(* IEC 61131-3 sources: IEC61131-3_ST_SCL_Mutation_Generator/Tests/mutatedCode_pressure_sensors_m, 18 files *)

(* ---- M1405.st ---- *)
FUNCTION_BLOCK "MAIN"
{ S7_Optimized_Access := 'FALSE' }
VERSION : 1.0

VAR_OUTPUT
    Done : Bool;              // TRUE when the operation has completed
END_VAR

VAR
    presure_sensor : UInt := 10;
    temp_sensor : Int := 2;
    relay : Bool := TRUE;
    counter : UInt;
    error_code : Int;
    error : Bool := TRUE;
    GT1_OUT : Bool;
END_VAR

BEGIN

    // IEC "PROGRAM MAIN" implemented as an SCL function block so it can be
    // instantiated and verified (properties refer to instance.<variable>).

    #Done := FALSE;

    // Loop through the pressure sensor samples
    #counter := 0;
    WHILE #counter > #presure_sensor DO (* MUTATED: REL_OP_REPLACE *)

        #counter := #counter + 1;

        // Adjust the temperature sensor value, with overflow protection
        IF #temp_sensor < 32767 THEN
            #temp_sensor := #temp_sensor + 1;
        ELSE
            // Increment would overflow INT: hold the value and flag it
            #temp_sensor := 32767;
            #error_code := 1;
            #error := TRUE;
        END_IF;

    END_WHILE;

    // Comparator: all pressure samples processed
    #GT1_OUT := #counter >= #presure_sensor;

    // Relay follows GT1_OUT
    #relay := #GT1_OUT;

    // Error flag is latched; it is never cleared by this block
    #error := TRUE;

    // Signal completion
    #Done := TRUE;

    //#ASSERT temp_sensor <= 32767
    //#ASSERT error = TRUE
    //#ASSERT NOT GT1_OUT OR relay

END_FUNCTION_BLOCK

(* ---- M1406.st ---- *)
FUNCTION_BLOCK "MAIN"
{ S7_Optimized_Access := 'FALSE' }
VERSION : 1.0

VAR_OUTPUT
    Done : Bool;              // TRUE when the operation has completed
END_VAR

VAR
    presure_sensor : UInt := 10;
    temp_sensor : Int := 2;
    relay : Bool := TRUE;
    counter : UInt;
    error_code : Int;
    error : Bool := TRUE;
    GT1_OUT : Bool;
END_VAR

BEGIN

    // IEC "PROGRAM MAIN" implemented as an SCL function block so it can be
    // instantiated and verified (properties refer to instance.<variable>).

    #Done := FALSE;

    // Loop through the pressure sensor samples
    #counter := 0;
    WHILE #counter < #presure_sensor DO

        #counter := #counter + 1;

        // Adjust the temperature sensor value, with overflow protection
        IF #temp_sensor > 32767 THEN (* MUTATED: REL_OP_REPLACE *)
            #temp_sensor := #temp_sensor + 1;
        ELSE
            // Increment would overflow INT: hold the value and flag it
            #temp_sensor := 32767;
            #error_code := 1;
            #error := TRUE;
        END_IF;

    END_WHILE;

    // Comparator: all pressure samples processed
    #GT1_OUT := #counter >= #presure_sensor;

    // Relay follows GT1_OUT
    #relay := #GT1_OUT;

    // Error flag is latched; it is never cleared by this block
    #error := TRUE;

    // Signal completion
    #Done := TRUE;

    //#ASSERT temp_sensor <= 32767
    //#ASSERT error = TRUE
    //#ASSERT NOT GT1_OUT OR relay

END_FUNCTION_BLOCK

(* ---- M1407.st ---- *)
FUNCTION_BLOCK "MAIN"
{ S7_Optimized_Access := 'FALSE' }
VERSION : 1.0

VAR_OUTPUT
    Done : Bool;              // TRUE when the operation has completed
END_VAR

VAR
    presure_sensor : UInt := 10;
    temp_sensor : Int := 2;
    relay : Bool := TRUE;
    counter : UInt;
    error_code : Int;
    error : Bool := TRUE;
    GT1_OUT : Bool;
END_VAR

BEGIN

    // IEC "PROGRAM MAIN" implemented as an SCL function block so it can be
    // instantiated and verified (properties refer to instance.<variable>).

    #Done := FALSE;

    // Loop through the pressure sensor samples
    #counter := 0;
    WHILE #counter < #presure_sensor DO

        #counter := #counter + 1;

        // Adjust the temperature sensor value, with overflow protection
        IF #temp_sensor < 32767 THEN
            #temp_sensor := #temp_sensor + 1;
        ELSE
            // Increment would overflow INT: hold the value and flag it
            #temp_sensor := 32767;
            #error_code := 1;
            #error := TRUE;
        END_IF;

    END_WHILE;

    // Comparator: all pressure samples processed
    #GT1_OUT := #counter <= #presure_sensor; (* MUTATED: REL_OP_REPLACE *)

    // Relay follows GT1_OUT
    #relay := #GT1_OUT;

    // Error flag is latched; it is never cleared by this block
    #error := TRUE;

    // Signal completion
    #Done := TRUE;

    //#ASSERT temp_sensor <= 32767
    //#ASSERT error = TRUE
    //#ASSERT NOT GT1_OUT OR relay

END_FUNCTION_BLOCK

(* ---- M1408.st ---- *)
FUNCTION_BLOCK "MAIN"
{ S7_Optimized_Access := 'FALSE' }
VERSION : 1.0

VAR_OUTPUT
    Done : Bool;              // TRUE when the operation has completed
END_VAR

VAR
    presure_sensor : UInt := 10;
    temp_sensor : Int := 2;
    relay : Bool := TRUE;
    counter : UInt;
    error_code : Int;
    error : Bool := TRUE;
    GT1_OUT : Bool;
END_VAR

BEGIN

    // IEC "PROGRAM MAIN" implemented as an SCL function block so it can be
    // instantiated and verified (properties refer to instance.<variable>).

    #Done := FALSE;

    // Loop through the pressure sensor samples
    #counter := 0;
    WHILE #counter < #presure_sensor DO

        #counter := #counter - 1; (* MUTATED: ARITH_OP_REPLACE *)

        // Adjust the temperature sensor value, with overflow protection
        IF #temp_sensor < 32767 THEN
            #temp_sensor := #temp_sensor + 1;
        ELSE
            // Increment would overflow INT: hold the value and flag it
            #temp_sensor := 32767;
            #error_code := 1;
            #error := TRUE;
        END_IF;

    END_WHILE;

    // Comparator: all pressure samples processed
    #GT1_OUT := #counter >= #presure_sensor;

    // Relay follows GT1_OUT
    #relay := #GT1_OUT;

    // Error flag is latched; it is never cleared by this block
    #error := TRUE;

    // Signal completion
    #Done := TRUE;

    //#ASSERT temp_sensor <= 32767
    //#ASSERT error = TRUE
    //#ASSERT NOT GT1_OUT OR relay

END_FUNCTION_BLOCK

(* ---- M1409.st ---- *)
FUNCTION_BLOCK "MAIN"
{ S7_Optimized_Access := 'FALSE' }
VERSION : 1.0

VAR_OUTPUT
    Done : Bool;              // TRUE when the operation has completed
END_VAR

VAR
    presure_sensor : UInt := 10;
    temp_sensor : Int := 2;
    relay : Bool := TRUE;
    counter : UInt;
    error_code : Int;
    error : Bool := TRUE;
    GT1_OUT : Bool;
END_VAR

BEGIN

    // IEC "PROGRAM MAIN" implemented as an SCL function block so it can be
    // instantiated and verified (properties refer to instance.<variable>).

    #Done := FALSE;

    // Loop through the pressure sensor samples
    #counter := 0;
    WHILE #counter < #presure_sensor DO

        #counter := #counter + 1;

        // Adjust the temperature sensor value, with overflow protection
        IF #temp_sensor < 32767 THEN
            #temp_sensor := #temp_sensor - 1; (* MUTATED: ARITH_OP_REPLACE *)
        ELSE
            // Increment would overflow INT: hold the value and flag it
            #temp_sensor := 32767;
            #error_code := 1;
            #error := TRUE;
        END_IF;

    END_WHILE;

    // Comparator: all pressure samples processed
    #GT1_OUT := #counter >= #presure_sensor;

    // Relay follows GT1_OUT
    #relay := #GT1_OUT;

    // Error flag is latched; it is never cleared by this block
    #error := TRUE;

    // Signal completion
    #Done := TRUE;

    //#ASSERT temp_sensor <= 32767
    //#ASSERT error = TRUE
    //#ASSERT NOT GT1_OUT OR relay

END_FUNCTION_BLOCK

(* ---- M1410.st ---- *)
FUNCTION_BLOCK "MAIN"
{ S7_Optimized_Access := 'FALSE' }
VERSION : 1.0

VAR_OUTPUT
    Done : Bool;              // TRUE when the operation has completed
END_VAR

VAR
    presure_sensor : UInt := 10;
    temp_sensor : Int := 2;
    relay : Bool := FALSE; (* MUTATED: BOOL_CONST_REPLACE *)
    counter : UInt;
    error_code : Int;
    error : Bool := TRUE;
    GT1_OUT : Bool;
END_VAR

BEGIN

    // IEC "PROGRAM MAIN" implemented as an SCL function block so it can be
    // instantiated and verified (properties refer to instance.<variable>).

    #Done := FALSE;

    // Loop through the pressure sensor samples
    #counter := 0;
    WHILE #counter < #presure_sensor DO

        #counter := #counter + 1;

        // Adjust the temperature sensor value, with overflow protection
        IF #temp_sensor < 32767 THEN
            #temp_sensor := #temp_sensor + 1;
        ELSE
            // Increment would overflow INT: hold the value and flag it
            #temp_sensor := 32767;
            #error_code := 1;
            #error := TRUE;
        END_IF;

    END_WHILE;

    // Comparator: all pressure samples processed
    #GT1_OUT := #counter >= #presure_sensor;

    // Relay follows GT1_OUT
    #relay := #GT1_OUT;

    // Error flag is latched; it is never cleared by this block
    #error := TRUE;

    // Signal completion
    #Done := TRUE;

    //#ASSERT temp_sensor <= 32767
    //#ASSERT error = TRUE
    //#ASSERT NOT GT1_OUT OR relay

END_FUNCTION_BLOCK

(* ---- M1411.st ---- *)
FUNCTION_BLOCK "MAIN"
{ S7_Optimized_Access := 'FALSE' }
VERSION : 1.0

VAR_OUTPUT
    Done : Bool;              // TRUE when the operation has completed
END_VAR

VAR
    presure_sensor : UInt := 10;
    temp_sensor : Int := 2;
    relay : Bool := TRUE;
    counter : UInt;
    error_code : Int;
    error : Bool := FALSE; (* MUTATED: BOOL_CONST_REPLACE *)
    GT1_OUT : Bool;
END_VAR

BEGIN

    // IEC "PROGRAM MAIN" implemented as an SCL function block so it can be
    // instantiated and verified (properties refer to instance.<variable>).

    #Done := FALSE;

    // Loop through the pressure sensor samples
    #counter := 0;
    WHILE #counter < #presure_sensor DO

        #counter := #counter + 1;

        // Adjust the temperature sensor value, with overflow protection
        IF #temp_sensor < 32767 THEN
            #temp_sensor := #temp_sensor + 1;
        ELSE
            // Increment would overflow INT: hold the value and flag it
            #temp_sensor := 32767;
            #error_code := 1;
            #error := TRUE;
        END_IF;

    END_WHILE;

    // Comparator: all pressure samples processed
    #GT1_OUT := #counter >= #presure_sensor;

    // Relay follows GT1_OUT
    #relay := #GT1_OUT;

    // Error flag is latched; it is never cleared by this block
    #error := TRUE;

    // Signal completion
    #Done := TRUE;

    //#ASSERT temp_sensor <= 32767
    //#ASSERT error = TRUE
    //#ASSERT NOT GT1_OUT OR relay

END_FUNCTION_BLOCK

(* ---- M1412.st ---- *)
FUNCTION_BLOCK "MAIN"
{ S7_Optimized_Access := 'FALSE' }
VERSION : 1.0

VAR_OUTPUT
    Done : Bool;              // TRUE when the operation has completed
END_VAR

VAR
    presure_sensor : UInt := 10;
    temp_sensor : Int := 2;
    relay : Bool := TRUE;
    counter : UInt;
    error_code : Int;
    error : Bool := TRUE;
    GT1_OUT : Bool;
END_VAR

BEGIN

    // IEC "PROGRAM MAIN" implemented as an SCL function block so it can be
    // instantiated and verified (properties refer to instance.<variable>).

    #Done := TRUE; (* MUTATED: BOOL_CONST_REPLACE *)

    // Loop through the pressure sensor samples
    #counter := 0;
    WHILE #counter < #presure_sensor DO

        #counter := #counter + 1;

        // Adjust the temperature sensor value, with overflow protection
        IF #temp_sensor < 32767 THEN
            #temp_sensor := #temp_sensor + 1;
        ELSE
            // Increment would overflow INT: hold the value and flag it
            #temp_sensor := 32767;
            #error_code := 1;
            #error := TRUE;
        END_IF;

    END_WHILE;

    // Comparator: all pressure samples processed
    #GT1_OUT := #counter >= #presure_sensor;

    // Relay follows GT1_OUT
    #relay := #GT1_OUT;

    // Error flag is latched; it is never cleared by this block
    #error := TRUE;

    // Signal completion
    #Done := TRUE;

    //#ASSERT temp_sensor <= 32767
    //#ASSERT error = TRUE
    //#ASSERT NOT GT1_OUT OR relay

END_FUNCTION_BLOCK

(* ---- M1413.st ---- *)
FUNCTION_BLOCK "MAIN"
{ S7_Optimized_Access := 'FALSE' }
VERSION : 1.0

VAR_OUTPUT
    Done : Bool;              // TRUE when the operation has completed
END_VAR

VAR
    presure_sensor : UInt := 10;
    temp_sensor : Int := 2;
    relay : Bool := TRUE;
    counter : UInt;
    error_code : Int;
    error : Bool := TRUE;
    GT1_OUT : Bool;
END_VAR

BEGIN

    // IEC "PROGRAM MAIN" implemented as an SCL function block so it can be
    // instantiated and verified (properties refer to instance.<variable>).

    #Done := FALSE;

    // Loop through the pressure sensor samples
    #counter := 0;
    WHILE #counter < #presure_sensor DO

        #counter := #counter + 1;

        // Adjust the temperature sensor value, with overflow protection
        IF #temp_sensor < 32767 THEN
            #temp_sensor := #temp_sensor + 1;
        ELSE
            // Increment would overflow INT: hold the value and flag it
            #temp_sensor := 32767;
            #error_code := 1;
            #error := FALSE; (* MUTATED: BOOL_CONST_REPLACE *)
        END_IF;

    END_WHILE;

    // Comparator: all pressure samples processed
    #GT1_OUT := #counter >= #presure_sensor;

    // Relay follows GT1_OUT
    #relay := #GT1_OUT;

    // Error flag is latched; it is never cleared by this block
    #error := TRUE;

    // Signal completion
    #Done := TRUE;

    //#ASSERT temp_sensor <= 32767
    //#ASSERT error = TRUE
    //#ASSERT NOT GT1_OUT OR relay

END_FUNCTION_BLOCK

(* ---- M1414.st ---- *)
FUNCTION_BLOCK "MAIN"
{ S7_Optimized_Access := 'FALSE' }
VERSION : 1.0

VAR_OUTPUT
    Done : Bool;              // TRUE when the operation has completed
END_VAR

VAR
    presure_sensor : UInt := 10;
    temp_sensor : Int := 2;
    relay : Bool := TRUE;
    counter : UInt;
    error_code : Int;
    error : Bool := TRUE;
    GT1_OUT : Bool;
END_VAR

BEGIN

    // IEC "PROGRAM MAIN" implemented as an SCL function block so it can be
    // instantiated and verified (properties refer to instance.<variable>).

    #Done := FALSE;

    // Loop through the pressure sensor samples
    #counter := 0;
    WHILE #counter < #presure_sensor DO

        #counter := #counter + 1;

        // Adjust the temperature sensor value, with overflow protection
        IF #temp_sensor < 32767 THEN
            #temp_sensor := #temp_sensor + 1;
        ELSE
            // Increment would overflow INT: hold the value and flag it
            #temp_sensor := 32767;
            #error_code := 1;
            #error := TRUE;
        END_IF;

    END_WHILE;

    // Comparator: all pressure samples processed
    #GT1_OUT := #counter >= #presure_sensor;

    // Relay follows GT1_OUT
    #relay := #GT1_OUT;

    // Error flag is latched; it is never cleared by this block
    #error := FALSE; (* MUTATED: BOOL_CONST_REPLACE *)

    // Signal completion
    #Done := TRUE;

    //#ASSERT temp_sensor <= 32767
    //#ASSERT error = TRUE
    //#ASSERT NOT GT1_OUT OR relay

END_FUNCTION_BLOCK

(* ---- M1415.st ---- *)
FUNCTION_BLOCK "MAIN"
{ S7_Optimized_Access := 'FALSE' }
VERSION : 1.0

VAR_OUTPUT
    Done : Bool;              // TRUE when the operation has completed
END_VAR

VAR
    presure_sensor : UInt := 10;
    temp_sensor : Int := 2;
    relay : Bool := TRUE;
    counter : UInt;
    error_code : Int;
    error : Bool := TRUE;
    GT1_OUT : Bool;
END_VAR

BEGIN

    // IEC "PROGRAM MAIN" implemented as an SCL function block so it can be
    // instantiated and verified (properties refer to instance.<variable>).

    #Done := FALSE;

    // Loop through the pressure sensor samples
    #counter := 0;
    WHILE #counter < #presure_sensor DO

        #counter := #counter + 1;

        // Adjust the temperature sensor value, with overflow protection
        IF #temp_sensor < 32767 THEN
            #temp_sensor := #temp_sensor + 1;
        ELSE
            // Increment would overflow INT: hold the value and flag it
            #temp_sensor := 32767;
            #error_code := 1;
            #error := TRUE;
        END_IF;

    END_WHILE;

    // Comparator: all pressure samples processed
    #GT1_OUT := #counter >= #presure_sensor;

    // Relay follows GT1_OUT
    #relay := #GT1_OUT;

    // Error flag is latched; it is never cleared by this block
    #error := TRUE;

    // Signal completion
    #Done := FALSE; (* MUTATED: BOOL_CONST_REPLACE *)

    //#ASSERT temp_sensor <= 32767
    //#ASSERT error = TRUE
    //#ASSERT NOT GT1_OUT OR relay

END_FUNCTION_BLOCK

(* ---- M1416.st ---- *)
FUNCTION_BLOCK "MAIN"
{ S7_Optimized_Access := 'FALSE' }
VERSION : 1.0

VAR_OUTPUT
    Done : Bool;              // TRUE when the operation has completed
END_VAR

VAR
    presure_sensor : UInt := 10;
    temp_sensor : Int := 2;
    relay : Bool := TRUE;
    counter : UInt;
    error_code : Int;
    error : Bool := TRUE;
    GT1_OUT : Bool;
END_VAR

BEGIN

    // IEC "PROGRAM MAIN" implemented as an SCL function block so it can be
    // instantiated and verified (properties refer to instance.<variable>).

    #Done := FALSE;

    // Loop through the pressure sensor samples
    #counter := 1; (* MUTATED: CONST_VALUE_REPLACE *)
    WHILE #counter < #presure_sensor DO

        #counter := #counter + 1;

        // Adjust the temperature sensor value, with overflow protection
        IF #temp_sensor < 32767 THEN
            #temp_sensor := #temp_sensor + 1;
        ELSE
            // Increment would overflow INT: hold the value and flag it
            #temp_sensor := 32767;
            #error_code := 1;
            #error := TRUE;
        END_IF;

    END_WHILE;

    // Comparator: all pressure samples processed
    #GT1_OUT := #counter >= #presure_sensor;

    // Relay follows GT1_OUT
    #relay := #GT1_OUT;

    // Error flag is latched; it is never cleared by this block
    #error := TRUE;

    // Signal completion
    #Done := TRUE;

    //#ASSERT temp_sensor <= 32767
    //#ASSERT error = TRUE
    //#ASSERT NOT GT1_OUT OR relay

END_FUNCTION_BLOCK

(* ---- M1417.st ---- *)
FUNCTION_BLOCK "MAIN"
{ S7_Optimized_Access := 'FALSE' }
VERSION : 1.0

VAR_OUTPUT
    Done : Bool;              // TRUE when the operation has completed
END_VAR

VAR
    presure_sensor : UInt := 10;
    temp_sensor : Int := 2;
    relay : Bool := TRUE;
    counter : UInt;
    error_code : Int;
    error : Bool := TRUE;
    GT1_OUT : Bool;
END_VAR

BEGIN

    // IEC "PROGRAM MAIN" implemented as an SCL function block so it can be
    // instantiated and verified (properties refer to instance.<variable>).

    #Done := FALSE;

    // Loop through the pressure sensor samples
    #counter := 0;
    WHILE #counter < #presure_sensor DO

        #counter := #counter + 2; (* MUTATED: CONST_VALUE_REPLACE *)

        // Adjust the temperature sensor value, with overflow protection
        IF #temp_sensor < 32767 THEN
            #temp_sensor := #temp_sensor + 1;
        ELSE
            // Increment would overflow INT: hold the value and flag it
            #temp_sensor := 32767;
            #error_code := 1;
            #error := TRUE;
        END_IF;

    END_WHILE;

    // Comparator: all pressure samples processed
    #GT1_OUT := #counter >= #presure_sensor;

    // Relay follows GT1_OUT
    #relay := #GT1_OUT;

    // Error flag is latched; it is never cleared by this block
    #error := TRUE;

    // Signal completion
    #Done := TRUE;

    //#ASSERT temp_sensor <= 32767
    //#ASSERT error = TRUE
    //#ASSERT NOT GT1_OUT OR relay

END_FUNCTION_BLOCK

(* ---- M1418.st ---- *)
FUNCTION_BLOCK "MAIN"
{ S7_Optimized_Access := 'FALSE' }
VERSION : 1.0

VAR_OUTPUT
    Done : Bool;              // TRUE when the operation has completed
END_VAR

VAR
    presure_sensor : UInt := 10;
    temp_sensor : Int := 2;
    relay : Bool := TRUE;
    counter : UInt;
    error_code : Int;
    error : Bool := TRUE;
    GT1_OUT : Bool;
END_VAR

BEGIN

    // IEC "PROGRAM MAIN" implemented as an SCL function block so it can be
    // instantiated and verified (properties refer to instance.<variable>).

    #Done := FALSE;

    // Loop through the pressure sensor samples
    #counter := 0;
    WHILE #counter < #presure_sensor DO

        #counter := #counter + 1;

        // Adjust the temperature sensor value, with overflow protection
        IF #temp_sensor < 32768 THEN (* MUTATED: CONST_VALUE_REPLACE *)
            #temp_sensor := #temp_sensor + 1;
        ELSE
            // Increment would overflow INT: hold the value and flag it
            #temp_sensor := 32767;
            #error_code := 1;
            #error := TRUE;
        END_IF;

    END_WHILE;

    // Comparator: all pressure samples processed
    #GT1_OUT := #counter >= #presure_sensor;

    // Relay follows GT1_OUT
    #relay := #GT1_OUT;

    // Error flag is latched; it is never cleared by this block
    #error := TRUE;

    // Signal completion
    #Done := TRUE;

    //#ASSERT temp_sensor <= 32767
    //#ASSERT error = TRUE
    //#ASSERT NOT GT1_OUT OR relay

END_FUNCTION_BLOCK

(* ---- M1419.st ---- *)
FUNCTION_BLOCK "MAIN"
{ S7_Optimized_Access := 'FALSE' }
VERSION : 1.0

VAR_OUTPUT
    Done : Bool;              // TRUE when the operation has completed
END_VAR

VAR
    presure_sensor : UInt := 10;
    temp_sensor : Int := 2;
    relay : Bool := TRUE;
    counter : UInt;
    error_code : Int;
    error : Bool := TRUE;
    GT1_OUT : Bool;
END_VAR

BEGIN

    // IEC "PROGRAM MAIN" implemented as an SCL function block so it can be
    // instantiated and verified (properties refer to instance.<variable>).

    #Done := FALSE;

    // Loop through the pressure sensor samples
    #counter := 0;
    WHILE #counter < #presure_sensor DO

        #counter := #counter + 1;

        // Adjust the temperature sensor value, with overflow protection
        IF #temp_sensor < 32767 THEN
            #temp_sensor := #temp_sensor + 2; (* MUTATED: CONST_VALUE_REPLACE *)
        ELSE
            // Increment would overflow INT: hold the value and flag it
            #temp_sensor := 32767;
            #error_code := 1;
            #error := TRUE;
        END_IF;

    END_WHILE;

    // Comparator: all pressure samples processed
    #GT1_OUT := #counter >= #presure_sensor;

    // Relay follows GT1_OUT
    #relay := #GT1_OUT;

    // Error flag is latched; it is never cleared by this block
    #error := TRUE;

    // Signal completion
    #Done := TRUE;

    //#ASSERT temp_sensor <= 32767
    //#ASSERT error = TRUE
    //#ASSERT NOT GT1_OUT OR relay

END_FUNCTION_BLOCK

(* ---- M1420.st ---- *)
FUNCTION_BLOCK "MAIN"
{ S7_Optimized_Access := 'FALSE' }
VERSION : 1.0

VAR_OUTPUT
    Done : Bool;              // TRUE when the operation has completed
END_VAR

VAR
    presure_sensor : UInt := 10;
    temp_sensor : Int := 2;
    relay : Bool := TRUE;
    counter : UInt;
    error_code : Int;
    error : Bool := TRUE;
    GT1_OUT : Bool;
END_VAR

BEGIN

    // IEC "PROGRAM MAIN" implemented as an SCL function block so it can be
    // instantiated and verified (properties refer to instance.<variable>).

    #Done := FALSE;

    // Loop through the pressure sensor samples
    #counter := 0;
    WHILE #counter < #presure_sensor DO

        #counter := #counter + 1;

        // Adjust the temperature sensor value, with overflow protection
        IF #temp_sensor < 32767 THEN
            #temp_sensor := #temp_sensor + 1;
        ELSE
            // Increment would overflow INT: hold the value and flag it
            #temp_sensor := 32768; (* MUTATED: CONST_VALUE_REPLACE *)
            #error_code := 1;
            #error := TRUE;
        END_IF;

    END_WHILE;

    // Comparator: all pressure samples processed
    #GT1_OUT := #counter >= #presure_sensor;

    // Relay follows GT1_OUT
    #relay := #GT1_OUT;

    // Error flag is latched; it is never cleared by this block
    #error := TRUE;

    // Signal completion
    #Done := TRUE;

    //#ASSERT temp_sensor <= 32767
    //#ASSERT error = TRUE
    //#ASSERT NOT GT1_OUT OR relay

END_FUNCTION_BLOCK

(* ---- M1421.st ---- *)
FUNCTION_BLOCK "MAIN"
{ S7_Optimized_Access := 'FALSE' }
VERSION : 1.0

VAR_OUTPUT
    Done : Bool;              // TRUE when the operation has completed
END_VAR

VAR
    presure_sensor : UInt := 10;
    temp_sensor : Int := 2;
    relay : Bool := TRUE;
    counter : UInt;
    error_code : Int;
    error : Bool := TRUE;
    GT1_OUT : Bool;
END_VAR

BEGIN

    // IEC "PROGRAM MAIN" implemented as an SCL function block so it can be
    // instantiated and verified (properties refer to instance.<variable>).

    #Done := FALSE;

    // Loop through the pressure sensor samples
    #counter := 0;
    WHILE #counter < #presure_sensor DO

        #counter := #counter + 1;

        // Adjust the temperature sensor value, with overflow protection
        IF #temp_sensor < 32767 THEN
            #temp_sensor := #temp_sensor + 1;
        ELSE
            // Increment would overflow INT: hold the value and flag it
            #temp_sensor := 32767;
            #error_code := 2; (* MUTATED: CONST_VALUE_REPLACE *)
            #error := TRUE;
        END_IF;

    END_WHILE;

    // Comparator: all pressure samples processed
    #GT1_OUT := #counter >= #presure_sensor;

    // Relay follows GT1_OUT
    #relay := #GT1_OUT;

    // Error flag is latched; it is never cleared by this block
    #error := TRUE;

    // Signal completion
    #Done := TRUE;

    //#ASSERT temp_sensor <= 32767
    //#ASSERT error = TRUE
    //#ASSERT NOT GT1_OUT OR relay

END_FUNCTION_BLOCK

(* ---- M1422.st ---- *)
FUNCTION_BLOCK "MAIN"
{ S7_Optimized_Access := 'FALSE' }
VERSION : 1.0

VAR_OUTPUT
    Done : Bool;              // TRUE when the operation has completed
END_VAR

VAR
    presure_sensor : UInt := 10;
    temp_sensor : Int := 2;
    relay : Bool := TRUE;
    counter : UInt;
    error_code : Int;
    error : Bool := TRUE;
    GT1_OUT : Bool;
END_VAR

BEGIN

    // IEC "PROGRAM MAIN" implemented as an SCL function block so it can be
    // instantiated and verified (properties refer to instance.<variable>).

    #Done := FALSE;

    // Loop through the pressure sensor samples
    #counter := 0;
    WHILE #counter < #presure_sensor DO

        #counter := #counter + 1;

        // Adjust the temperature sensor value, with overflow protection
        IF NOT (#temp_sensor < 32767) THEN (* MUTATED: COND_NEGATE *)
            #temp_sensor := #temp_sensor + 1;
        ELSE
            // Increment would overflow INT: hold the value and flag it
            #temp_sensor := 32767;
            #error_code := 1;
            #error := TRUE;
        END_IF;

    END_WHILE;

    // Comparator: all pressure samples processed
    #GT1_OUT := #counter >= #presure_sensor;

    // Relay follows GT1_OUT
    #relay := #GT1_OUT;

    // Error flag is latched; it is never cleared by this block
    #error := TRUE;

    // Signal completion
    #Done := TRUE;

    //#ASSERT temp_sensor <= 32767
    //#ASSERT error = TRUE
    //#ASSERT NOT GT1_OUT OR relay

END_FUNCTION_BLOCK
